{attribute 'TcGvlVarFlags' := 'OPC'}
VAR_GLOBAL
    // I/O module state — Python can read inputs and write output setpoints
    // ADS symbol: GVL_IO.stIO
    stIO            : ST_IOData;
END_VAR

(* stored: Version 1.1.0.1, ProductVersion 3.1.4026.18
   GVL GVL_IO: Id {b73b097a-b8d4-49fc-aa49-e2f6a25c0235} *)
